// SIMATIC S7-200 project (STEP 7-Micro/WIN), CPU 224 CN REL 02.01

SYMBOL_TABLE USUARIO1
SM1              I0.0     // Detecta el vàstago extendidio del pistòn pequeño
SM2              I0.1     // Detecta el vàstago retraido del piston pequeño
SM3              I0.2     // Detecta el vastago extendido del piston largo
SM4              I0.3     // Detecta el vastago retraido del piston largo
SF1              I0.4     // Detecta la presencia de una pieza en el final de la unidad de alimentacion
SF2              I0.5     // Detecta la presencia de pieza en la parte superior del cilindro
SF3              I0.6     // Detecta la presencia de pieza en la parte inferior del cilindro
SI1              I0.7     // Detecta la presencia de una pieza metàlica en la parte inferior del cilindro
SV1              I1.2     // Boton de inicio
SR1              I1.3     // Boton disponible para su uso
QS               I1.4     // Detiene el proceso en cualquier instante de tiempo
SA               I1.5     // Switch disponible para su uso
KM1              Q0.0     // Acciona la electrovaluvula que controla el piston pequeño
KM2              Q0.1     // Acciona la electrovalvula
HL1              Q0.7     // Lampara disponible (Anomalia y precaucion)
HL2              Q1.0     // Lampara disponible (Funcionamiento normal)
HL3              Q1.1     // Lampara disponible (Emergencia y peligro)
END_SYMBOL_TABLE

ORGANIZATION_BLOCK PRINCIPAL:OB1
TITLE=UNIDAD DE ALIMENTACIÒN
BEGIN
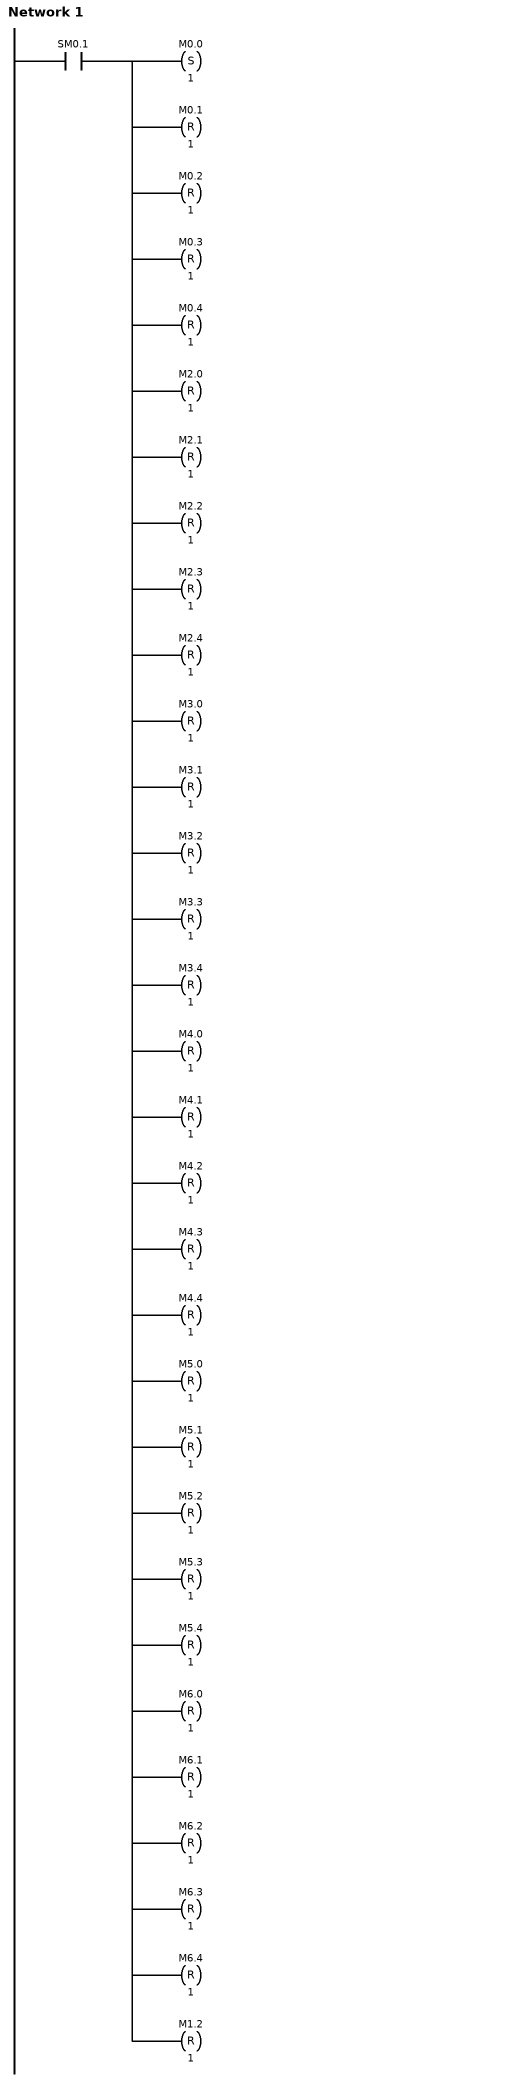
Network 1
LD     SM0.1
S      M0.0, 1
R      M0.1, 1
R      M0.2, 1
R      M0.3, 1
R      M0.4, 1
R      M2.0, 1
R      M2.1, 1
R      M2.2, 1
R      M2.3, 1
R      M2.4, 1
R      M3.0, 1
R      M3.1, 1
R      M3.2, 1
R      M3.3, 1
R      M3.4, 1
R      M4.0, 1
R      M4.1, 1
R      M4.2, 1
R      M4.3, 1
R      M4.4, 1
R      M5.0, 1
R      M5.1, 1
R      M5.2, 1
R      M5.3, 1
R      M5.4, 1
R      M6.0, 1
R      M6.1, 1
R      M6.2, 1
R      M6.3, 1
R      M6.4, 1
R      M1.2, 1
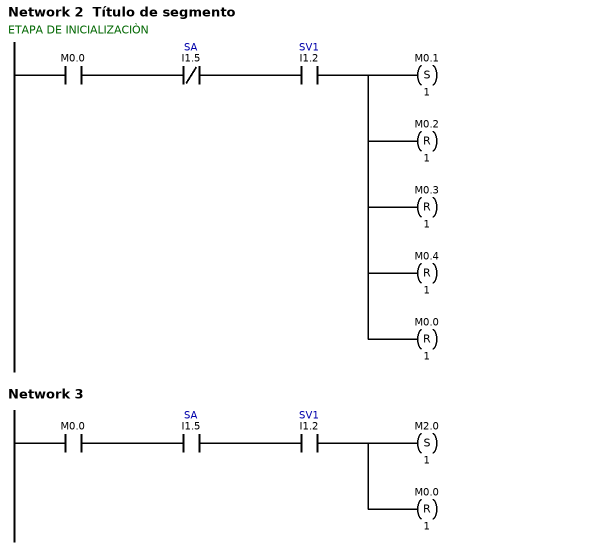
Network 2 // Título de segmento
// ETAPA DE INICIALIZACIÒN
LD     M0.0
AN     SA:I1.5
A      SV1:I1.2
S      M0.1, 1
R      M0.2, 1
R      M0.3, 1
R      M0.4, 1
R      M0.0, 1
Network 3
LD     M0.0
A      SA:I1.5
A      SV1:I1.2
S      M2.0, 1
R      M0.0, 1
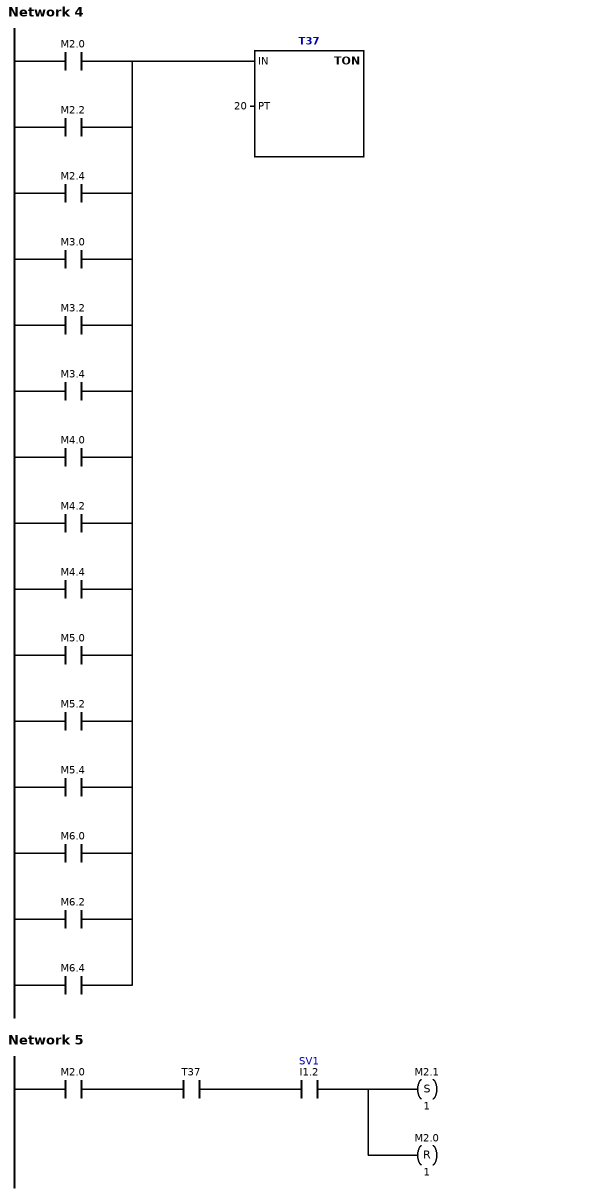
Network 4
LD     M2.0
O      M2.2
O      M2.4
O      M3.0
O      M3.2
O      M3.4
O      M4.0
O      M4.2
O      M4.4
O      M5.0
O      M5.2
O      M5.4
O      M6.0
O      M6.2
O      M6.4
TON    T37, 20
Network 5
LD     M2.0
A      T37
A      SV1:I1.2
S      M2.1, 1
R      M2.0, 1
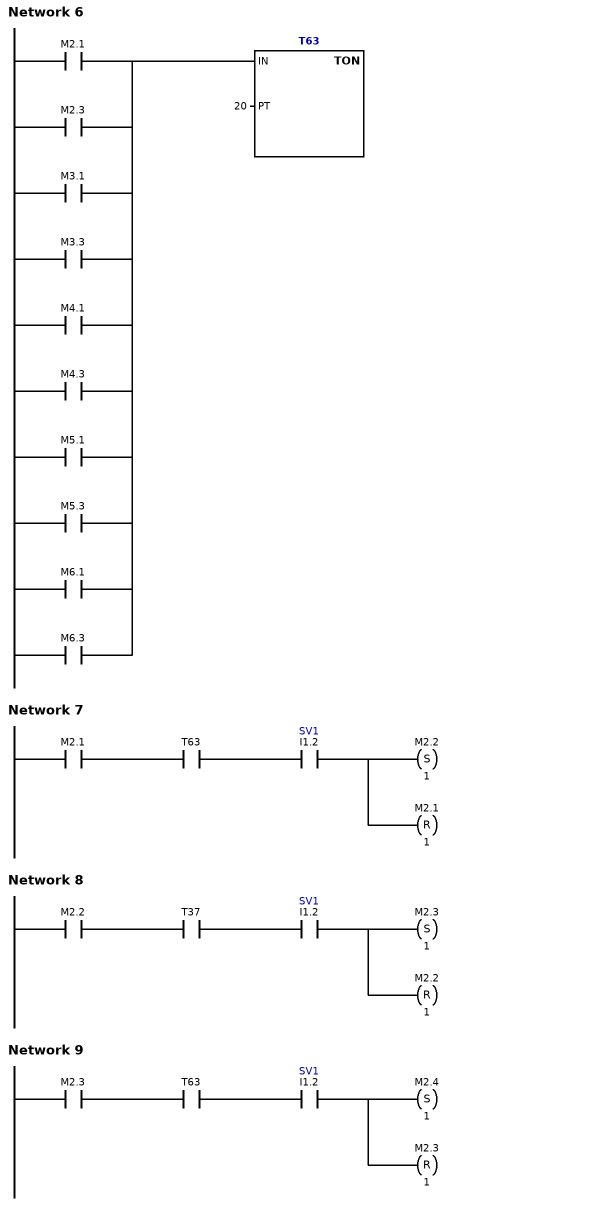
Network 6
LD     M2.1
O      M2.3
O      M3.1
O      M3.3
O      M4.1
O      M4.3
O      M5.1
O      M5.3
O      M6.1
O      M6.3
TON    T63, 20
Network 7
LD     M2.1
A      T63
A      SV1:I1.2
S      M2.2, 1
R      M2.1, 1
Network 8
LD     M2.2
A      T37
A      SV1:I1.2
S      M2.3, 1
R      M2.2, 1
Network 9
LD     M2.3
A      T63
A      SV1:I1.2
S      M2.4, 1
R      M2.3, 1
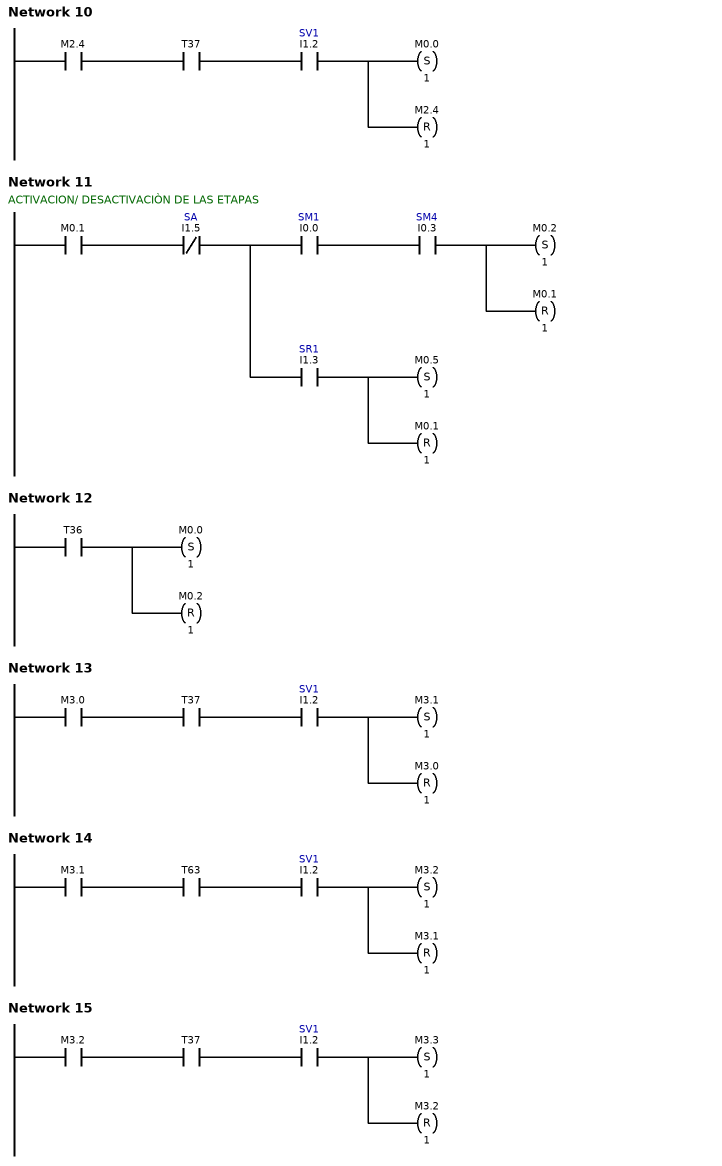
Network 10
LD     M2.4
A      T37
A      SV1:I1.2
S      M0.0, 1
R      M2.4, 1
Network 11
// ACTIVACION/ DESACTIVACIÒN DE LAS ETAPAS
LD     M0.1
AN     SA:I1.5
LPS
A      SM1:I0.0
A      SM4:I0.3
S      M0.2, 1
R      M0.1, 1
LPP
A      SR1:I1.3
S      M0.5, 1
R      M0.1, 1
Network 12
LD     T36
S      M0.0, 1
R      M0.2, 1
Network 13
LD     M3.0
A      T37
A      SV1:I1.2
S      M3.1, 1
R      M3.0, 1
Network 14
LD     M3.1
A      T63
A      SV1:I1.2
S      M3.2, 1
R      M3.1, 1
Network 15
LD     M3.2
A      T37
A      SV1:I1.2
S      M3.3, 1
R      M3.2, 1
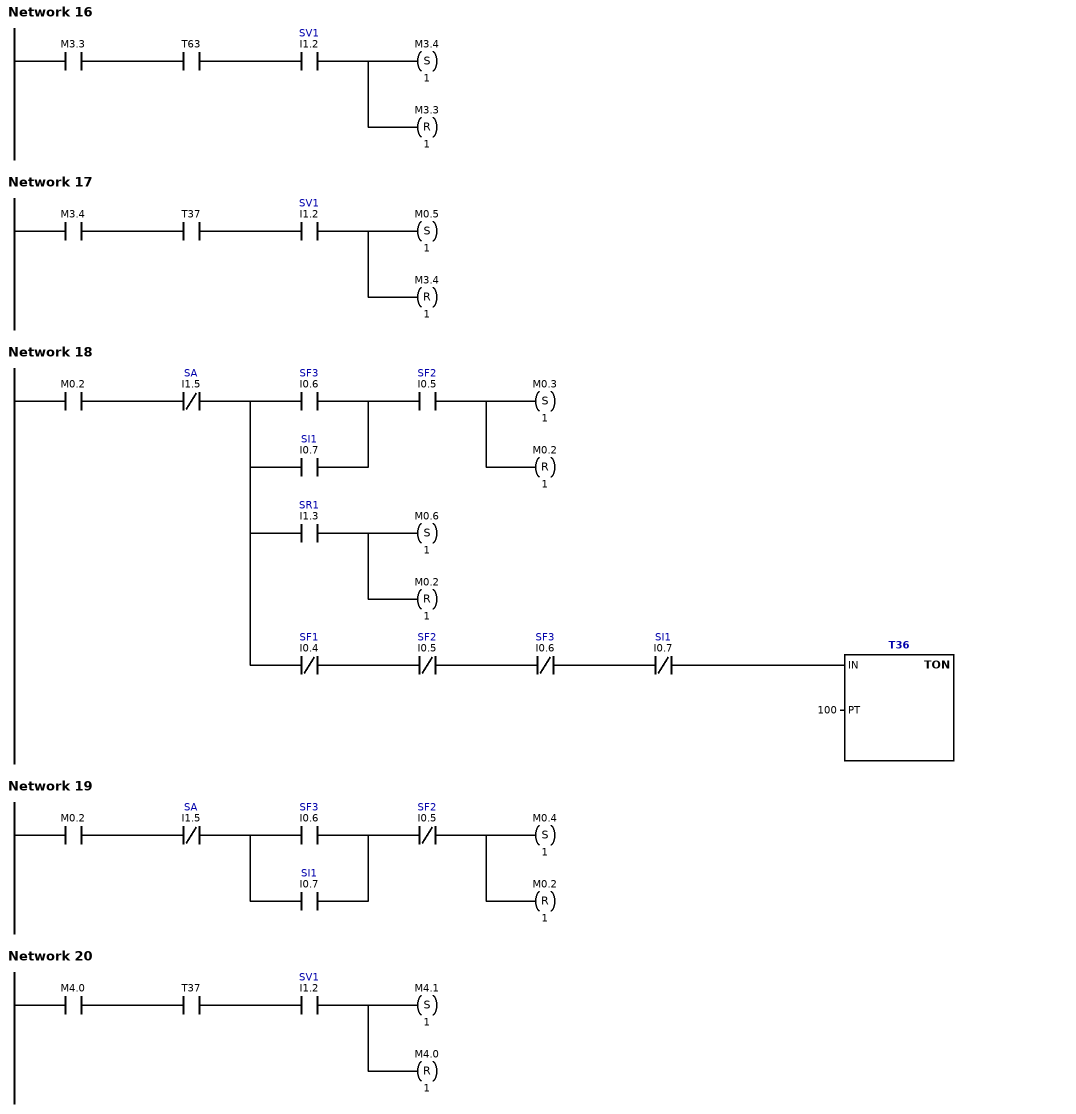
Network 16
LD     M3.3
A      T63
A      SV1:I1.2
S      M3.4, 1
R      M3.3, 1
Network 17
LD     M3.4
A      T37
A      SV1:I1.2
S      M0.5, 1
R      M3.4, 1
Network 18
LD     M0.2
AN     SA:I1.5
LPS
LD     SF3:I0.6
O      SI1:I0.7
A      SF2:I0.5
ALD
S      M0.3, 1
R      M0.2, 1
LRD
A      SR1:I1.3
S      M0.6, 1
R      M0.2, 1
LPP
AN     SF1:I0.4
AN     SF2:I0.5
AN     SF3:I0.6
AN     SI1:I0.7
TON    T36, 100
Network 19
LD     M0.2
AN     SA:I1.5
LD     SF3:I0.6
O      SI1:I0.7
ALD
AN     SF2:I0.5
S      M0.4, 1
R      M0.2, 1
Network 20
LD     M4.0
A      T37
A      SV1:I1.2
S      M4.1, 1
R      M4.0, 1
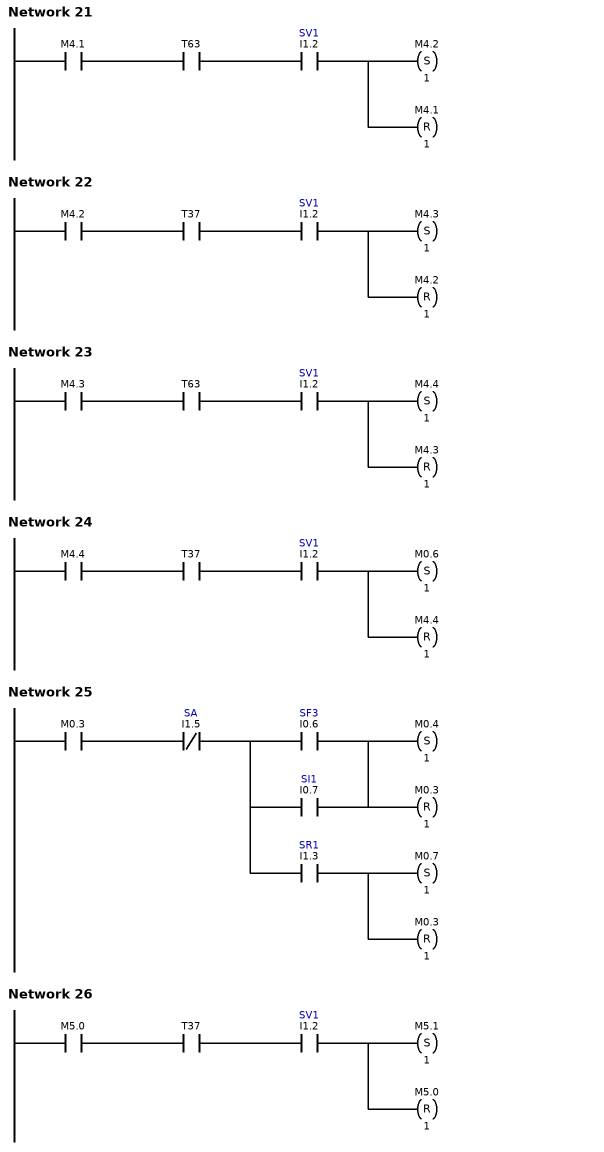
Network 21
LD     M4.1
A      T63
A      SV1:I1.2
S      M4.2, 1
R      M4.1, 1
Network 22
LD     M4.2
A      T37
A      SV1:I1.2
S      M4.3, 1
R      M4.2, 1
Network 23
LD     M4.3
A      T63
A      SV1:I1.2
S      M4.4, 1
R      M4.3, 1
Network 24
LD     M4.4
A      T37
A      SV1:I1.2
S      M0.6, 1
R      M4.4, 1
Network 25
LD     M0.3
AN     SA:I1.5
LPS
LD     SF3:I0.6
O      SI1:I0.7
ALD
S      M0.4, 1
R      M0.3, 1
LPP
A      SR1:I1.3
S      M0.7, 1
R      M0.3, 1
Network 26
LD     M5.0
A      T37
A      SV1:I1.2
S      M5.1, 1
R      M5.0, 1
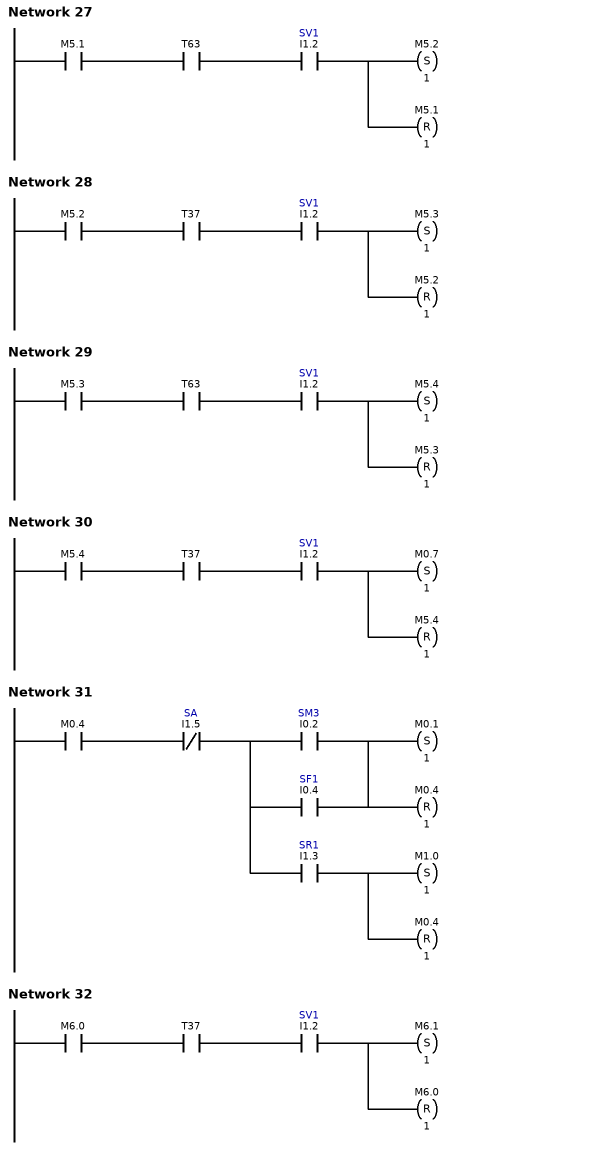
Network 27
LD     M5.1
A      T63
A      SV1:I1.2
S      M5.2, 1
R      M5.1, 1
Network 28
LD     M5.2
A      T37
A      SV1:I1.2
S      M5.3, 1
R      M5.2, 1
Network 29
LD     M5.3
A      T63
A      SV1:I1.2
S      M5.4, 1
R      M5.3, 1
Network 30
LD     M5.4
A      T37
A      SV1:I1.2
S      M0.7, 1
R      M5.4, 1
Network 31
LD     M0.4
AN     SA:I1.5
LPS
LD     SM3:I0.2
O      SF1:I0.4
ALD
S      M0.1, 1
R      M0.4, 1
LPP
A      SR1:I1.3
S      M1.0, 1
R      M0.4, 1
Network 32
LD     M6.0
A      T37
A      SV1:I1.2
S      M6.1, 1
R      M6.0, 1
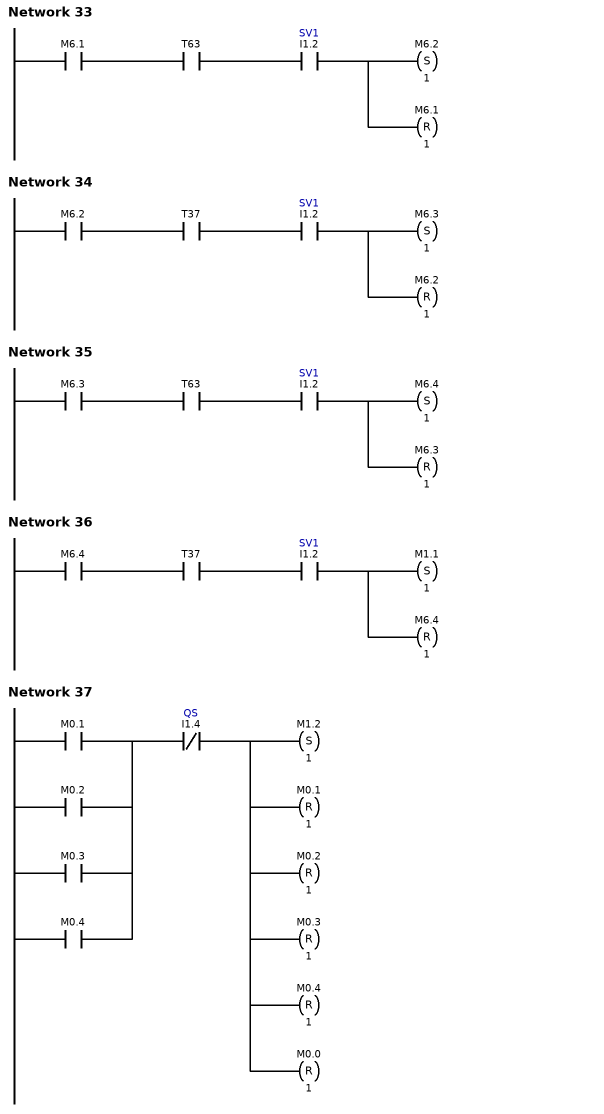
Network 33
LD     M6.1
A      T63
A      SV1:I1.2
S      M6.2, 1
R      M6.1, 1
Network 34
LD     M6.2
A      T37
A      SV1:I1.2
S      M6.3, 1
R      M6.2, 1
Network 35
LD     M6.3
A      T63
A      SV1:I1.2
S      M6.4, 1
R      M6.3, 1
Network 36
LD     M6.4
A      T37
A      SV1:I1.2
S      M1.1, 1
R      M6.4, 1
Network 37
LD     M0.1
O      M0.2
O      M0.3
O      M0.4
AN     QS:I1.4
S      M1.2, 1
R      M0.1, 1
R      M0.2, 1
R      M0.3, 1
R      M0.4, 1
R      M0.0, 1
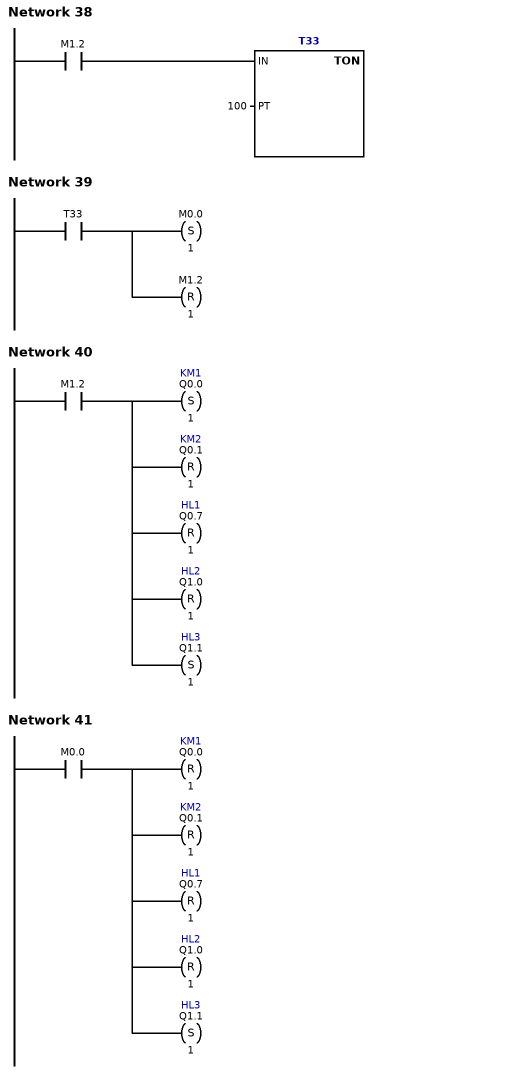
Network 38
LD     M1.2
TON    T33, 100
Network 39
LD     T33
S      M0.0, 1
R      M1.2, 1
Network 40
LD     M1.2
S      KM1:Q0.0, 1
R      KM2:Q0.1, 1
R      HL1:Q0.7, 1
R      HL2:Q1.0, 1
S      HL3:Q1.1, 1
Network 41
LD     M0.0
R      KM1:Q0.0, 1
R      KM2:Q0.1, 1
R      HL1:Q0.7, 1
R      HL2:Q1.0, 1
S      HL3:Q1.1, 1
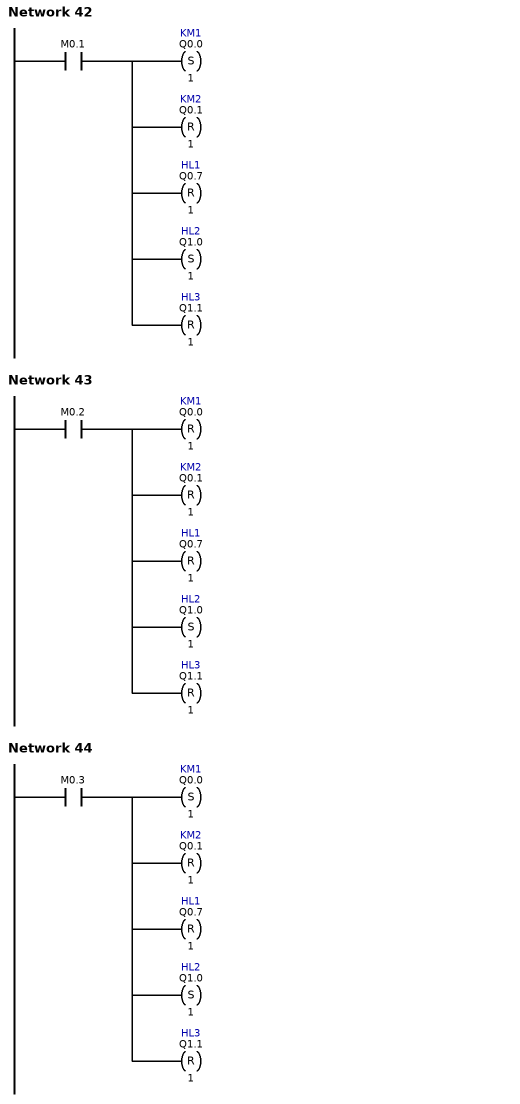
Network 42
LD     M0.1
S      KM1:Q0.0, 1
R      KM2:Q0.1, 1
R      HL1:Q0.7, 1
S      HL2:Q1.0, 1
R      HL3:Q1.1, 1
Network 43
LD     M0.2
R      KM1:Q0.0, 1
R      KM2:Q0.1, 1
R      HL1:Q0.7, 1
S      HL2:Q1.0, 1
R      HL3:Q1.1, 1
Network 44
LD     M0.3
S      KM1:Q0.0, 1
R      KM2:Q0.1, 1
R      HL1:Q0.7, 1
S      HL2:Q1.0, 1
R      HL3:Q1.1, 1
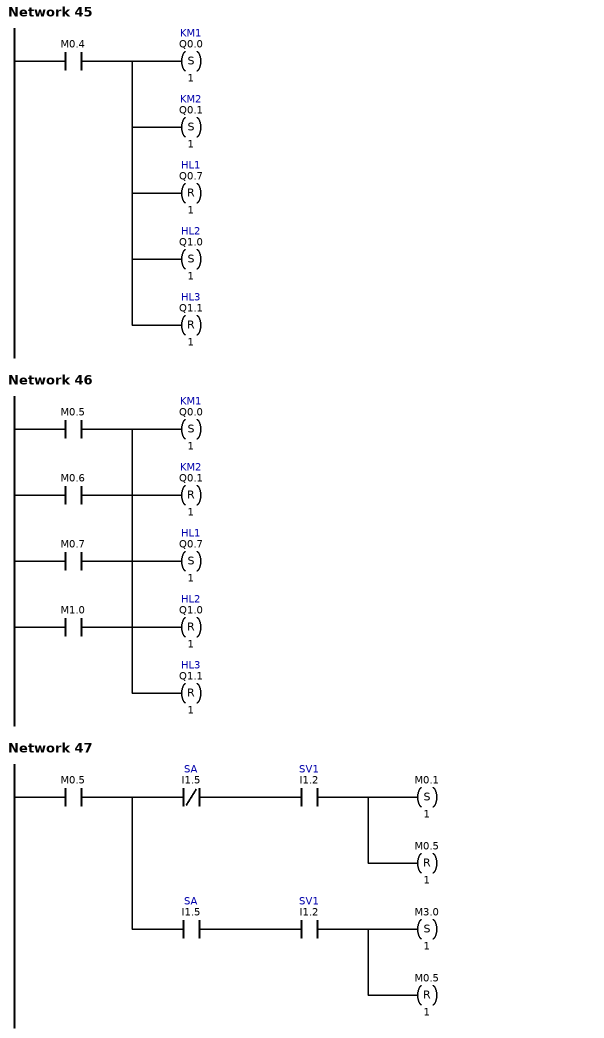
Network 45
LD     M0.4
S      KM1:Q0.0, 1
S      KM2:Q0.1, 1
R      HL1:Q0.7, 1
S      HL2:Q1.0, 1
R      HL3:Q1.1, 1
Network 46
LD     M0.5
O      M0.6
O      M0.7
O      M1.0
S      KM1:Q0.0, 1
R      KM2:Q0.1, 1
S      HL1:Q0.7, 1
R      HL2:Q1.0, 1
R      HL3:Q1.1, 1
Network 47
LD     M0.5
LPS
AN     SA:I1.5
A      SV1:I1.2
S      M0.1, 1
R      M0.5, 1
LPP
A      SA:I1.5
A      SV1:I1.2
S      M3.0, 1
R      M0.5, 1
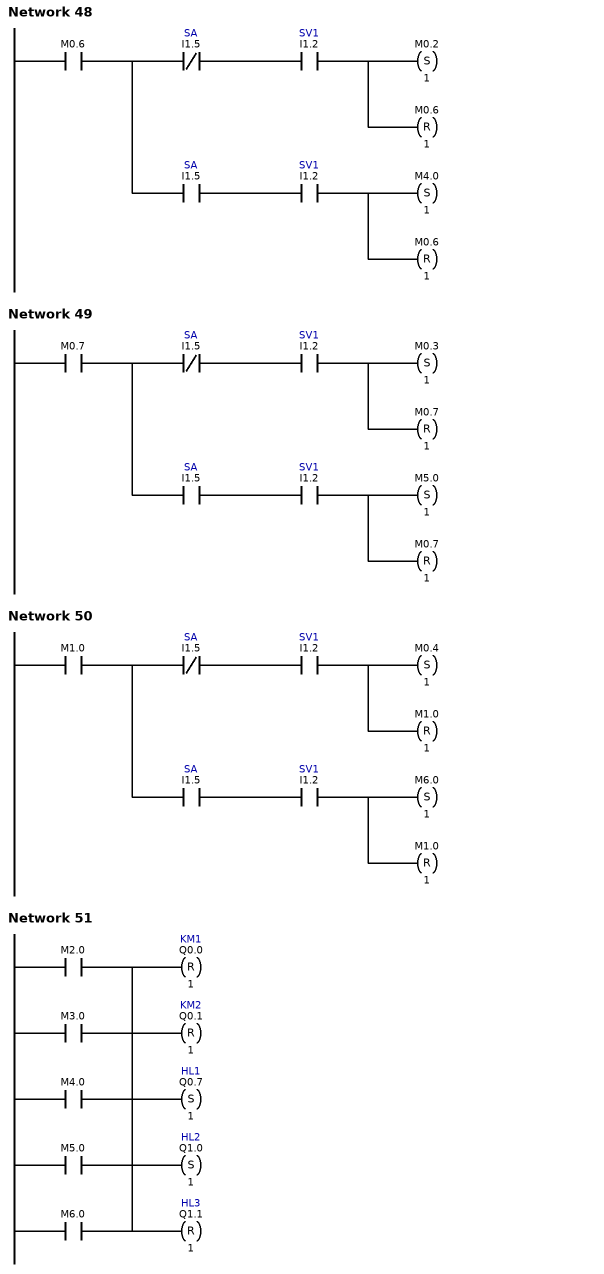
Network 48
LD     M0.6
LPS
AN     SA:I1.5
A      SV1:I1.2
S      M0.2, 1
R      M0.6, 1
LPP
A      SA:I1.5
A      SV1:I1.2
S      M4.0, 1
R      M0.6, 1
Network 49
LD     M0.7
LPS
AN     SA:I1.5
A      SV1:I1.2
S      M0.3, 1
R      M0.7, 1
LPP
A      SA:I1.5
A      SV1:I1.2
S      M5.0, 1
R      M0.7, 1
Network 50
LD     M1.0
LPS
AN     SA:I1.5
A      SV1:I1.2
S      M0.4, 1
R      M1.0, 1
LPP
A      SA:I1.5
A      SV1:I1.2
S      M6.0, 1
R      M1.0, 1
Network 51
LD     M2.0
O      M3.0
O      M4.0
O      M5.0
O      M6.0
R      KM1:Q0.0, 1
R      KM2:Q0.1, 1
S      HL1:Q0.7, 1
S      HL2:Q1.0, 1
R      HL3:Q1.1, 1
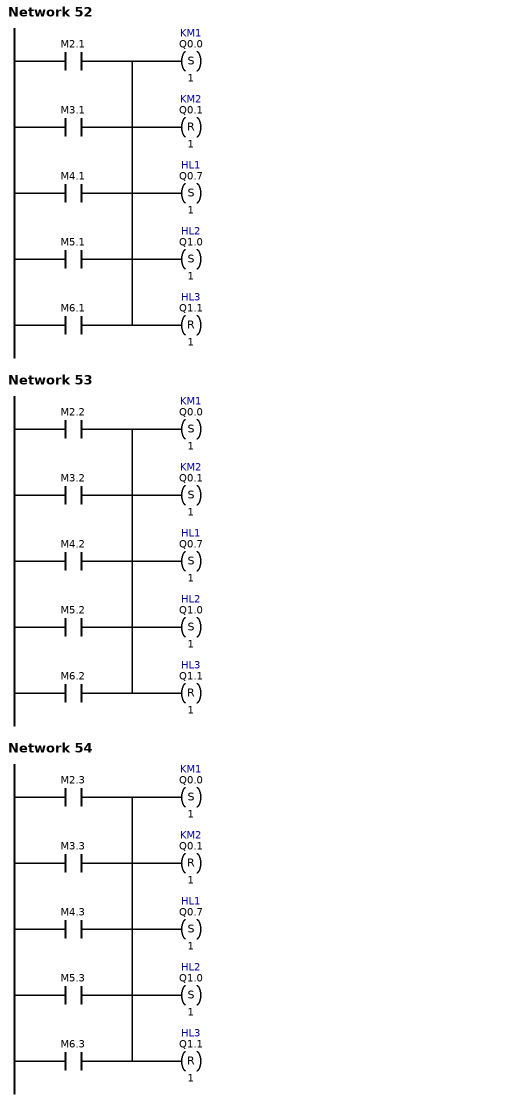
Network 52
LD     M2.1
O      M3.1
O      M4.1
O      M5.1
O      M6.1
S      KM1:Q0.0, 1
R      KM2:Q0.1, 1
S      HL1:Q0.7, 1
S      HL2:Q1.0, 1
R      HL3:Q1.1, 1
Network 53
LD     M2.2
O      M3.2
O      M4.2
O      M5.2
O      M6.2
S      KM1:Q0.0, 1
S      KM2:Q0.1, 1
S      HL1:Q0.7, 1
S      HL2:Q1.0, 1
R      HL3:Q1.1, 1
Network 54
LD     M2.3
O      M3.3
O      M4.3
O      M5.3
O      M6.3
S      KM1:Q0.0, 1
R      KM2:Q0.1, 1
S      HL1:Q0.7, 1
S      HL2:Q1.0, 1
R      HL3:Q1.1, 1
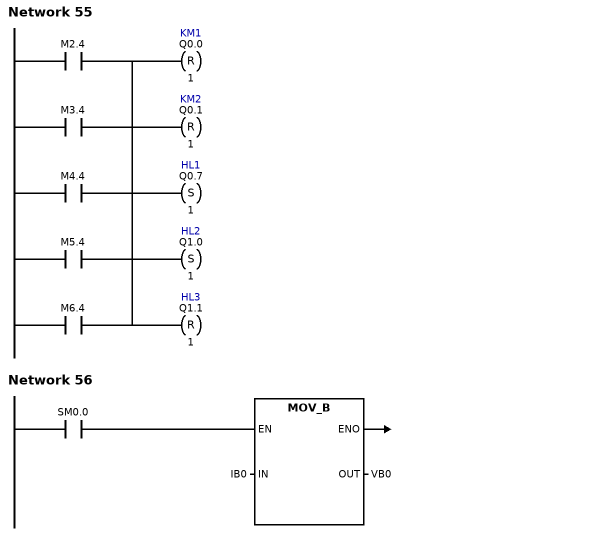
Network 55
LD     M2.4
O      M3.4
O      M4.4
O      M5.4
O      M6.4
R      KM1:Q0.0, 1
R      KM2:Q0.1, 1
S      HL1:Q0.7, 1
S      HL2:Q1.0, 1
R      HL3:Q1.1, 1
Network 56
LD     SM0.0
MOVB   IB0, VB0
END_ORGANIZATION_BLOCK
